(* IEC 61131-3 sources: plcassist-cli/packages/volt-lsp-iec/test-corpus/lenze-mid/Device/Plc Logic/Application/Library Manager/VisuUserManagement, 50 files *)

(* ---- GVL_USERMGMTPROVIDER.gvl ---- *)
VAR_GLOBAL
	G_ARRUSERSTODISPLAY : ARRAY [0..14] OF VUM_UserInternal;
END_VAR

(* ---- VUM_ERRORCODES.gvl ---- *)
VAR_GLOBAL
	ERR_OK : UDINT := 16#0;
	ERR_FAILED : UDINT := 16#1;
	ERR_PARAMETER : UDINT := 16#2;
	ERR_VUM_FILE_NOT_FOUND : UDINT := 16#5000;
	ERR_VUM_TEMP_FILE_CANNOT_BE_OPENED : UDINT := 16#5001;
	ERR_VUM_FILE_READ_FAILED : UDINT := 16#5002;
	ERR_VUM_FILE_WRITE_FAILED : UDINT := 16#5003;
	ERR_VUM_INVALID_FILE_CONTENT : UDINT := 16#5004;
	ERR_VUM_USERNAME_ALREADY_EXIST : UDINT := 16#5005;
	ERR_VUM_WRONG_PASSWORD : UDINT := 16#5006;
	ERR_VUM_UNEQUAL_PASSWORD : UDINT := 16#5007;
	ERR_VUM_NEW_USER_DB_CANNOT_BE_STORED : UDINT := 16#5008;
	ERR_VUM_ONLY_VISIBLE_USERS_CAN_BE_REMOVED : UDINT := 16#5009;
	ERR_VUM_EMPTY_PASSWORD_NOT_ALLOWED : UDINT := 16#500A;
	ERR_VUM_ANOTHER_CLIENT_EDITS_UM : UDINT := 16#500B;
	ERR_VUM_SYSFILE_ERROR : UDINT := 16#500C;
	ERR_VUM_SETNEWUSERDB_FAILED : UDINT := 16#500D;
	ERR_VUM_PROXY_IS_NOT_IN_IDLE_MODE : UDINT := 16#500E;
	ERR_VUM_DATASERVER_ERROR : UDINT := 16#500F;
	ERR_VUM_DATASERVER_ERROR_USERS : UDINT := 16#5010;
	ERR_VUM_MAX_GROUP_LIMIT : UDINT := 16#5011;
	ERR_VUM_USER_DOES_NOT_EXIST : UDINT := 16#5012;
	ERR_VUM_USER_IS_INACTIVE : UDINT := 16#5013;
	ERR_VUM_NO_LOGIN_PROVIDER_AVAILABLE : UDINT := 16#5014;
	ERR_VUM_NO_CLIENT_MEMORY : UDINT := 16#5015;
	ERR_VUM_NO_USER_LOGGED_IN : UDINT := 16#5016;
	ERR_VUM_NO_VALID_USERGROUP_SET : UDINT := 16#5017;
	ERR_VUM_NO_RIGHT_TO_CHANGE_USERS : UDINT := 16#5018;
	ERR_VUM_NO_USER_MANAGEMENT : UDINT := 16#5019;
	ERR_VUM_USER_NOT_IN_USER_GROUP : UDINT := 16#501A;
	ERR_VUM_EXTERNAL_USER_DATABASE_PROVIDER2_NOT_IMPLEMENTED : UDINT := 16#501B;
	ERR_VUM_LOGIN_WRONG_ATTEMPT : UDINT := 16#501C;
	ERR_VUM_LOGIN_SECONDLAST_WRONG_ATTEMPT : UDINT := 16#501D;
	ERR_VUM_LOGIN_LOCKOUT_TEMP : UDINT := 16#501E;
	ERR_VUM_LOGIN_LOCKOUT_COMPLETE : UDINT := 16#501F;
	ERR_VUM_EMPTY_USER_NAME_NOT_ALLOWED : UDINT := 16#5020;
END_VAR

(* ---- VUM_EVENTS.gvl ---- *)
VAR_GLOBAL
	EVT_VISUUSERMGMTGETUSERCOUNT : UDINT := 16#10001;
	EVT_VISUUSERMGMTGETUSERS : UDINT := 16#10002;
	EVT_VISUUSERMGMTCHECKCHANGEUSER : UDINT := 16#10003;
	EVT_VISUUSERMGMTGETSETDB : UDINT := 16#10004;
	CMPID_CMPVISUSERVER : DWORD := 16#57;
END_VAR

(* ---- VUM_GVL.gvl ---- *)
VAR_GLOBAL
	G_VISUUSERMGMT : IVisuUserManagement4;
	G_VISUUSERMGMT2 : IVisuUserManagement4;
	G_VISUUSERMGMTINTERN : IVisuUserMgmt;
	G_STAPPLICATIONNAME : STRING := '';
	G_VUMUSERGROUPNAMES : ARRAY [0..MAX_USER_GROUPS] OF WSTRING;
	G_VUMUSERGROUPMAXINDEX : DWORD;
	G_BUSEVISUUSERMGMTDATASERVER : BOOL;
	G_UDILASTERROR : UDINT;
	G_SILOGINMAXATTEMPTS : SINT := -1;
	G_ILOGINLOCKOUTTIME : INT := -1;
	G_LOGINMAXATTEMPTSENTRIES : VisuUserMgmtFbLoginMaxAttemptsInfoVector;
	G_LOGINLOCKOUTENTRIES : VisuUserMgmtFbLoginLockoutTimeInfoVector;
	G_VISUUSERMANAGERCOMPONENT : STRING := 'VisuUserManager';
	G_VISUUSERMGMTLOGINDIALOGNAME : STRING := 'VUM_Login';
	G_VISUUSERMGMTCHANGEPASSWORDDIALOGNAME : STRING := 'VUM_ChangePassword';
	G_VISUUSERMGMTUSERMANAGEMENTDIALOGNAME : STRING := 'VisuUserManagement.VUM_UserManagementWide';
	G_VISUUSERMGMTRTSBASED : BOOL := FALSE;
	G_VISUUSERMGMTRTSBASEDPATHNAME : WSTRING(256) := "";
END_VAR

(* ---- VUM_GVL_CONSTANT.gvl ---- *)
VAR_GLOBAL
	USERGROUPFLAG_RIGHT_TO_CHANGE_USER : DWORD := 16#1;
	OUTPUT_INFO : INT := 16#1;
	OUTPUT_WARNING : INT := 16#2;
	OUTPUT_ERROR : INT := 16#4;
	OUTPUT_DEBUG : INT := 16#10;
	INVALID_USERGROUP_ID : DWORD := 16#FFFFFFFF;
	INVALID_DB_ID : DWORD := 16#FFFFFFFF;
	INVALID_SELECTION_OR_POS : DWORD := 16#FFFFFFFF;
	COMMENT_CHAR : WORD := 16#23;
	MAX_VISIBLE_USERS : UDINT := 3;
	MAX_USER_GROUPS : UDINT := 255;
	VISU_USER_MGMT_VERSION : DWORD := 0;
	GETSETDB_FLAGS_GETDB : UINT := 16#1;
	GETSETDB_FLAGS_SETDB : UINT := 16#2;
	GETSETDB_FLAGS_SET_RESULT_OK : UINT := 16#4;
	CHECKCHANGEUSER_FLAGS_CHECKLOGIN : UINT := 16#1;
	CHECKCHANGEUSER_FLAGS_CHANGEUSER : UINT := 16#2;
	INVALID_HANDLE : DWORD := 16#FFFFFFFF;
	TIMER_VALUE_LOCKOUT_ADMIN_USER : SINT := 10;
END_VAR

(* ---- VUM_GVL_PROVIDER.gvl ---- *)
VAR_GLOBAL
	G_VISUUSERMGMTPROVIDER : VisuUserMgmtProvider;
	G_BVISUUSERMGMTDIALOGOPEN : BOOL := FALSE;
	G_POPENUSERMGMTORPASSWORDCLIENT : POINTER TO VisuElems.VisuStructClientData;
	G_VISUCHANGEPASSWORDPROVIDER : VisuChangePasswordProvider;
	G_BVISUCHANGEPASSWORDDIALOGOPEN : BOOL := FALSE;
	G_VISUCHANGEPASSWORDPROVIDERMANAGER : Visu_FbChangePasswordProviderManager;
	G_VISULOGINPROVIDERMANAGER : Visu_FbLoginProviderManager;
END_VAR

(* ---- VUM_GVL_RTSUSERMGT.gvl ---- *)
VAR_GLOBAL
	ASSIGNRTSBASEDUSERMGT : VisuAssignRtsBasedUserMgt;
END_VAR

(* ---- IVISUUSERMGMT.itf ---- *)
INTERFACE IVISUUSERMGMT
END_INTERFACE

METHOD CHANGEUSER : BOOL
VAR_INPUT
	DWUSERDB : DWORD;
	PVUMUSER : POINTER TO VUM_User;
	UDIINDEX : UDINT;
	EEDITTYPE : VUM_EditType;
END_VAR
END_METHOD

METHOD CHANGEUSERPASSWORD : BOOL
VAR_INPUT
	DWUSERDB : DWORD;
	WSTUSERNAME : WSTRING;
	WSTNEWPASSWORD : WSTRING;
	WSTOLDPASSWORD : WSTRING;
END_VAR
END_METHOD

METHOD CHECKLOGININTERN : UDINT
VAR_INPUT
	WSTUSERNAME : WSTRING;
	WSTPASSWORD : WSTRING;
END_VAR
VAR_OUTPUT
	WSTFULLNAME : WSTRING;
	DWUSERGROUPID : DWORD;
END_VAR
END_METHOD

METHOD FILLLANGUAGEGROUPNAMES : BOOL
END_METHOD

METHOD GETCURRENTUSER : VUM_User
END_METHOD

METHOD GETGROUPCOUNT : DWORD
END_METHOD

METHOD GETGROUPFROMID : POINTER TO VUM_UserGroup
VAR_INPUT
	DWGROUPID : DWORD;
END_VAR
END_METHOD

METHOD GETGROUPIDFROMINDEX : DWORD
VAR_INPUT
	UDIINDEX : DWORD;
END_VAR
END_METHOD

METHOD GETGROUPINDEXFROMID : DWORD
VAR_INPUT
	DWGROUPID : DWORD;
END_VAR
END_METHOD

METHOD GETLASTERROR : UDINT
END_METHOD

METHOD GETTEXTIDFROMGROUPID : DWORD
VAR_INPUT
	DWGROUPID : DWORD;
END_VAR
END_METHOD

METHOD GETUSERCOUNT : UDINT
VAR_INPUT
	DWUSERDB : DWORD;
END_VAR
END_METHOD

METHOD GETUSERDBASCOPY : DWORD
END_METHOD

METHOD GETUSERS : DWORD
VAR_INPUT
	DWUSERDB : DWORD;
	UDISTARTINDEX : UDINT;
	UDIENDINDEX : UDINT;
	PARR : POINTER TO ARRAY [0..0] OF VUM_User;
	UDIARRSIZE : UDINT;
END_VAR
END_METHOD

METHOD REGISTEREXTERNALUSERDATABASEPROVIDER : VUM_ReturnValues
VAR_INPUT
	ITFEXTENALUSERDATABASEPROVIDER : IExternalUserDatabaseProvider;
END_VAR
END_METHOD

METHOD SETLASTERROR : BOOL
VAR_INPUT
	UDILASTERROR : UDINT;
END_VAR
END_METHOD

METHOD SETNEWUSERDB : BOOL
VAR_INPUT
	DWUSERDB : DWORD;
	BRESULTOK : BOOL;
END_VAR
END_METHOD

METHOD SETPROVIDER : BOOL
VAR_INPUT
	ITFVISUUSERMGMTPROVIDER : IVisuUserMgmtProvider;
END_VAR
END_METHOD

(* ---- IVISUUSERMGMT2.itf ---- *)
INTERFACE IVISUUSERMGMT2
END_INTERFACE

METHOD CHECKTEMPORARYLOCKEDUSER : BOOL
END_METHOD

(* ---- IVISUUSERMGMT3.itf ---- *)
INTERFACE IVISUUSERMGMT3
END_INTERFACE

METHOD CHANGEUSER3 : BOOL
VAR_INPUT
	PCLIENTDATA : POINTER TO VisuElems.VisuStructClientData;
	DWUSERDB : DWORD;
	PVUMUSERNEW : POINTER TO VUM_User;
	PVUMUSEROLD : POINTER TO VUM_User;
	UDIINDEX : UDINT;
	EEDITTYPE : VUM_EditType;
END_VAR
END_METHOD

METHOD CHANGEUSERPASSWORD3 : UDINT
VAR_INPUT
	PCLIENTDATA : POINTER TO VisuElems.VisuStructClientData;
	DWUSERDB : DWORD;
	WSTUSERNAME : WSTRING;
	WSTNEWPASSWORD : WSTRING;
	WSTOLDPASSWORD : WSTRING;
END_VAR
END_METHOD

METHOD CHECKADMINRIGHTS : VUM_UserAdminAccess
VAR_INPUT
	PCLIENTDATA : POINTER TO VisuElems.VisuStructClientData;
END_VAR
END_METHOD

METHOD CHECKGROUPS : BOOL
VAR_INPUT
	PCLIENTDATA : POINTER TO VisuElems.VisuStructClientData;
END_VAR
END_METHOD

METHOD GETUSERCOUNT3 : UDINT
VAR_INPUT
	PCLIENTDATA : POINTER TO VisuElems.VisuStructClientData;
	DWUSERDB : DWORD;
END_VAR
VAR_OUTPUT
	RESULT : RTS_IEC_RESULT;
END_VAR
END_METHOD

METHOD GETUSERS3 : DWORD
VAR_INPUT
	PCLIENTDATA : POINTER TO VisuElems.VisuStructClientData;
	DWUSERDB : DWORD;
	UDISTARTINDEX : UDINT;
	UDIENDINDEX : UDINT;
	PARR : POINTER TO ARRAY [0..0] OF VUM_User;
	UDIARRSIZE : UDINT;
END_VAR
END_METHOD

METHOD LOGINRTS : UDINT
VAR_INPUT
	WSTUSERNAME : WSTRING;
	WSTPASSWORD : WSTRING;
	PCLIENTDATA : POINTER TO VisuElems.VisuStructClientData;
	PUSER : POINTER TO VUM_User;
END_VAR
VAR_OUTPUT
	WSTFULLNAME : WSTRING;
	DWUSERGROUPID : DWORD;
END_VAR
END_METHOD

(* ---- IVISUUSERMGMT4.itf ---- *)
INTERFACE IVISUUSERMGMT4
END_INTERFACE

METHOD CHANGEUSER4 : BOOL
VAR_INPUT
	PCLIENTDATA : POINTER TO VisuElems.VisuStructClientData;
	DWUSERDB : DWORD;
	PVUMUSERNEW : POINTER TO VUM_UserInternal;
	PVUMUSEROLD : POINTER TO VUM_UserInternal;
	UDIINDEX : UDINT;
	EEDITTYPE : VUM_EditType;
END_VAR
END_METHOD

METHOD GETUSERS4 : DWORD
VAR_INPUT
	PCLIENTDATA : POINTER TO VisuElems.VisuStructClientData;
	DWUSERDB : DWORD;
	UDISTARTINDEX : UDINT;
	UDIENDINDEX : UDINT;
	PARR : POINTER TO ARRAY [0..0] OF VUM_UserInternal;
	UDIARRSIZE : UDINT;
END_VAR
END_METHOD

METHOD LOGOUTRTS
VAR_INPUT
	PCLIENTDATA : POINTER TO VisuElems.VisuStructClientData;
END_VAR
END_METHOD

(* ---- IVISUUSERMGMTPROVIDER.itf ---- *)
INTERFACE IVISUUSERMGMTPROVIDER
END_INTERFACE

METHOD SETUSERCOUNT : BOOL
VAR_INPUT
	UDIUSERCOUNT : UDINT;
END_VAR
END_METHOD

METHOD SETUSERDB : BOOL
VAR_INPUT
	UDIUSERDB : UDINT;
END_VAR
END_METHOD

METHOD SETUSERS : BOOL
VAR_INPUT
	UDIUSERCOUNT : UDINT;
	PARRUSERS : POINTER TO ARRAY [0..(MAX_VISIBLE_USERS - 1)] OF VUM_User;
END_VAR
END_METHOD

(* ---- COPYVUM_USER.fun ---- *)
FUNCTION COPYVUM_USER : BOOL
VAR_INPUT
	PVUM_USER : POINTER TO VUM_User;
	PVUM_USERINTERNAL : POINTER TO VUM_UserInternal;
	XFROMUSERTOINTERNAL : BOOL;
END_VAR
END_FUNCTION

(* ---- COPYVUM_USER3.fun ---- *)
FUNCTION COPYVUM_USER3 : BOOL
VAR_INPUT
	PVUM_USER3 : POINTER TO VUM_User3;
	PVUM_USERINTERNAL : POINTER TO VUM_UserInternal;
	XFROMUSERTOINTERNAL : BOOL;
END_VAR
END_FUNCTION

(* ---- FILTERERRORCODE.fun ---- *)
FUNCTION FILTERERRORCODE : UDINT
VAR_INPUT
	ERROR : UDINT;
END_VAR
END_FUNCTION

(* ---- HASUSERGROUPADMINRIGHTS.fun ---- *)
FUNCTION HASUSERGROUPADMINRIGHTS : BOOL
VAR_INPUT
	PUSERGROUP : POINTER TO VUM_UserGroup;
	PCLIENTDATA : POINTER TO VisuElems.VisuStructClientData;
END_VAR
END_FUNCTION

(* ---- ONCHANGEPASSWORDDIALOGCLOSED.fun ---- *)
FUNCTION ONCHANGEPASSWORDDIALOGCLOSED : BOOL
VAR_INPUT
	PCLIENTDATA : POINTER TO VisuElems.VisuStructClientData;
END_VAR
END_FUNCTION

(* ---- ONLOGINDIALOGCLOSED.fun ---- *)
FUNCTION ONLOGINDIALOGCLOSED : BOOL
VAR_INPUT
	PCLIENTDATA : POINTER TO VisuElems.VisuStructClientData;
END_VAR
END_FUNCTION

(* ---- ONUSERMANAGEMENTDIALOGCLOSED.fun ---- *)
FUNCTION ONUSERMANAGEMENTDIALOGCLOSED : BOOL
VAR_INPUT
	PCLIENTDATA : POINTER TO VisuElems.VisuStructClientData;
END_VAR
END_FUNCTION

(* ---- OPENCHANGEPASSWORDDIALOG.fun ---- *)
FUNCTION OPENCHANGEPASSWORDDIALOG : BOOL
VAR_INPUT
	PCLIENTDATA : POINTER TO VisuElems.VisuStructClientData;
END_VAR
END_FUNCTION

(* ---- OPENLOGINDIALOG.fun ---- *)
FUNCTION OPENLOGINDIALOG : BOOL
VAR_INPUT
	PCLIENTDATA : POINTER TO VisuElems.VisuStructClientData;
END_VAR
END_FUNCTION

(* ---- OPENUSERMANAGEMENTDIALOG.fun ---- *)
FUNCTION OPENUSERMANAGEMENTDIALOG : BOOL
VAR_INPUT
	PCLIENTDATA : POINTER TO VisuElems.VisuStructClientData;
END_VAR
END_FUNCTION

(* ---- PRVCHECKUSERMGRISACTIVE.fun ---- *)
FUNCTION PRVCHECKUSERMGRISACTIVE : BOOL
END_FUNCTION

(* ---- SWAPBYTEARRAYBYWORDS.fun ---- *)
FUNCTION SWAPBYTEARRAYBYWORDS : BOOL
VAR_INPUT
	PDATA : POINTER TO ARRAY [0..20] OF BYTE;
	DWSIZE : DWORD;
END_VAR
END_FUNCTION

(* ---- UTILFILLLANGUAGEGROUPNAMES.fun ---- *)
FUNCTION UTILFILLLANGUAGEGROUPNAMES : BOOL
VAR_INPUT
	PARRUSERGROUPTEXTIDS : POINTER TO ARRAY [0..0] OF DWORD;
	DWARRAYSIZE : DWORD;
END_VAR
END_FUNCTION

(* ---- UTILGETFILESIZE.fun ---- *)
FUNCTION UTILGETFILESIZE : UDINT
VAR_INPUT
	DWHANDLE : SysFile.RTS_IEC_HANDLE;
	STFILENAME : REFERENCE TO STRING(255);
	PULRESULT : POINTER TO UDINT;
END_VAR
END_FUNCTION

(* ---- UTILGETMD5HASH.fun ---- *)
FUNCTION UTILGETMD5HASH : BOOL
VAR_INPUT
	PDATA : POINTER TO BYTE;
	DWSIZE : DWORD;
	PMD5HASH : POINTER TO ARRAY [0..15] OF BYTE;
	BADDMAGICNUMBER : BOOL;
	BBYTEORDERMOTOROLAONPOWERPC : BOOL;
END_VAR
END_FUNCTION

(* ---- VISU_FCTINTELBYTEORDER.fun ---- *)
FUNCTION VISU_FCTINTELBYTEORDER : BOOL
END_FUNCTION

(* ---- VISUCREATEUSERMGMTOBJECTS.fun ---- *)
FUNCTION VISUCREATEUSERMGMTOBJECTS : RTS_IEC_RESULT
VAR_INPUT
	PUSERGROUPS : POINTER TO ARRAY [0..0] OF VUM_UserGroup;
	IARRAYSIZE : INT;
	PSAPPNAME : POINTER TO WSTRING;
END_VAR
END_FUNCTION

(* ---- VISUUSERMGMTHASUSERRIGHTTOCHANGEUSERS.fun ---- *)
FUNCTION VISUUSERMGMTHASUSERRIGHTTOCHANGEUSERS : BOOL
VAR_INPUT
	PVUMUSER : POINTER TO VUM_User;
	ITFVISUUSERMGMT : IVisuUserMgmt;
END_VAR
END_FUNCTION

(* ---- VISUUSERMGMTISRTS_GE_35_8.fun ---- *)
FUNCTION VISUUSERMGMTISRTS_GE_35_8 : BOOL
END_FUNCTION

(* ---- VISUUSERMGMTLOG.fun ---- *)
FUNCTION VISUUSERMGMTLOG : BOOL
VAR_INPUT
	DICLASS : DINT;
	DIERROR : DINT;
	DIINFO : DINT;
	STMESSAGE : STRING(255);
END_VAR
END_FUNCTION

(* ---- VISUUSERMGMTSERIALIZEVERSION.fun ---- *)
FUNCTION VISUUSERMGMTSERIALIZEVERSION : DWORD
VAR_INPUT
	VER : VERSION;
END_VAR
END_FUNCTION

(* ---- GLOBALTEXTLIST.fb ---- *)
FUNCTION_BLOCK GLOBALTEXTLIST
VAR
	M_TEXTLISTFILE : STRING(255);
	_STNAMESPACE : STRING;
END_VAR
END_FUNCTION_BLOCK

(* ---- IMAGEPOOL.fb ---- *)
FUNCTION_BLOCK IMAGEPOOL
VAR
	M_STNAMESPACE : STRING(80);
	M_STHELPVARID : STRING;
	M_STHELPVARPATH : STRING(255);
	M_STHELP : STRING;
	M_REGISTERIMAGES : BOOL := TRUE;
END_VAR
END_FUNCTION_BLOCK

METHOD FB_INIT : BOOL
VAR_INPUT
	BINITRETAINS : BOOL;
	BINCOPYCODE : BOOL;
END_VAR
END_METHOD

METHOD FB_REINIT : BOOL
END_METHOD

METHOD FB_EXIT : BOOL
VAR_INPUT
	BINCOPYCODE : BOOL;
END_VAR
END_METHOD

(* ---- IP_VUM.fb ---- *)
FUNCTION_BLOCK IP_VUM
VAR
	M_STNAMESPACE : STRING(80);
	M_STHELPVARID : STRING;
	M_STHELPVARPATH : STRING(255);
	M_STHELP : STRING;
	M_REGISTERIMAGES : BOOL := TRUE;
END_VAR
END_FUNCTION_BLOCK

METHOD FB_INIT : BOOL
VAR_INPUT
	BINITRETAINS : BOOL;
	BINCOPYCODE : BOOL;
END_VAR
END_METHOD

METHOD FB_REINIT : BOOL
END_METHOD

METHOD FB_EXIT : BOOL
VAR_INPUT
	BINCOPYCODE : BOOL;
END_VAR
END_METHOD

(* ---- TL_VUM_ERRORS.fb ---- *)
FUNCTION_BLOCK TL_VUM_ERRORS
VAR
	M_TEXTLISTFILE : STRING(255);
	_STNAMESPACE : STRING;
END_VAR
END_FUNCTION_BLOCK

(* ---- VISU_FBCHANGEPASSWORDPROVIDERMANAGER.fb ---- *)
FUNCTION_BLOCK VISU_FBCHANGEPASSWORDPROVIDERMANAGER
VAR
	M_ARRPROVIDER : ARRAY [0..(MAX_PROVIDER - 1)] OF VisuChangePasswordProvider;
	M_ARRCLIENT : ARRAY [0..(MAX_PROVIDER - 1)] OF POINTER TO VisuElems.VisuStructClientData;
	M_ITFCLIENTMANAGERLISTENER : VisuElems.IClientManagerListener := THIS^;
	M_BINIT : BOOL;
	I : INT;
	MAX_PROVIDER : INT := 5;
END_VAR
END_FUNCTION_BLOCK

METHOD FB_EXIT : BOOL
VAR_INPUT
	BINCOPYCODE : BOOL;
END_VAR
END_METHOD

METHOD INITIALIZE : BOOL
END_METHOD

METHOD REGISTERCLIENT : POINTER TO VisuChangePasswordProvider
VAR_INPUT
	PCLIENTDATA : POINTER TO VisuElems.VisuStructClientData;
END_VAR
END_METHOD

METHOD UNREGISTERCLIENT : BOOL
VAR_INPUT
	PCLIENTDATA : POINTER TO VisuElems.VisuStructClientData;
END_VAR
END_METHOD

METHOD CLIENTCREATED
VAR_INPUT
	PCLIENTDATA : POINTER TO VisuElems.VisuStructClientData;
END_VAR
END_METHOD

METHOD CLIENTDESTROYED
VAR_INPUT
	PCLIENTDATA : POINTER TO VisuElems.VisuStructClientData;
END_VAR
END_METHOD

(* ---- VISU_FBLOGINPROVIDERMANAGER.fb ---- *)
FUNCTION_BLOCK VISU_FBLOGINPROVIDERMANAGER
VAR
	M_ARRLOGINPROVIDER : ARRAY [0..(MAX_LOGIN_PROVIDER - 1)] OF VisuLoginProvider;
	M_ARRLOGINPROVIDERSET : ARRAY [0..(MAX_LOGIN_PROVIDER - 1)] OF BOOL;
	M_ITFCLIENTMANAGERLISTENER : VisuElems.IClientManagerListener := THIS^;
	M_BINIT : BOOL;
	I : INT;
	MAX_LOGIN_PROVIDER : INT := 5;
END_VAR
END_FUNCTION_BLOCK

METHOD FB_EXIT : BOOL
VAR_INPUT
	BINCOPYCODE : BOOL;
END_VAR
END_METHOD

METHOD INITIALIZE : BOOL
END_METHOD

METHOD REGISTERLOGINPROVIDERCLIENT : POINTER TO VisuLoginProvider
VAR_INPUT
	PCLIENTDATA : POINTER TO VisuElems.VisuStructClientData;
END_VAR
END_METHOD

METHOD UNREGISTERLOGINPROVIDERCLIENT : BOOL
VAR_INPUT
	PCLIENTDATA : POINTER TO VisuElems.VisuStructClientData;
END_VAR
END_METHOD

METHOD CLIENTCREATED
VAR_INPUT
	PCLIENTDATA : POINTER TO VisuElems.VisuStructClientData;
END_VAR
END_METHOD

METHOD CLIENTDESTROYED
VAR_INPUT
	PCLIENTDATA : POINTER TO VisuElems.VisuStructClientData;
END_VAR
END_METHOD

(* ---- VISUASSIGNRTSBASEDUSERMGT.fb ---- *)
FUNCTION_BLOCK VISUASSIGNRTSBASEDUSERMGT
VAR
	XSTATUSVISUUSERMGMTRTSBASED : BOOL;
END_VAR
END_FUNCTION_BLOCK

METHOD FB_EXIT : BOOL
VAR_INPUT
	BINCOPYCODE : BOOL;
END_VAR
END_METHOD

METHOD FB_INIT : BOOL
VAR_INPUT
	BINITRETAINS : BOOL;
	BINCOPYCODE : BOOL;
END_VAR
END_METHOD

(* ---- VISUCHANGEPASSWORDPROVIDER.fb ---- *)
FUNCTION_BLOCK VISUCHANGEPASSWORDPROVIDER
VAR
	STUSERNAME : WSTRING;
	STOLDPASSWORD : WSTRING;
	STPASSWORD : WSTRING;
	WSTOLDPASSWORD : WSTRING;
	STACKNOWLEDGEPASSWORD : WSTRING;
	DWDIALOGRESULTOK : BOOL;
	DWLASTDIALOGRESULTOK : BOOL;
	DWDIALOGRESULTCANCEL : BOOL;
	DWLASTDIALOGRESULTCANCEL : BOOL;
	UDILASTERROR : UDINT;
	DWRESULT : DWORD;
	VUMUSER : VUM_User;
	BRTSBASED : BOOL;
	BCHGPASSWORD : BOOL;
	_IVISUUSERMGMT : IVisuUserMgmt;
	_IVISUUSERMGMT4 : IVisuUserMgmt4;
	_VISUUSERMGMTSTATE : EVisuUserMgmtState;
	_PCLIENTDATA : POINTER TO VisuElems.VisuStructClientData;
	_BCURRENTSTATE : BYTE := 0;
	_BLASTCURRENTSTATE : BYTE := 0;
	_DWUSERDB : DWORD;
	VCPP_STATE_NONE : BYTE := 0;
	VCPP_STATE_GET_USER_DB : BYTE := 1;
	VCPP_STATE_CHECK_LOGIN : BYTE := 2;
	VCPP_STATE_CHANGE_USER_PASSWORD : BYTE := 3;
	VCPP_STATE_SET_USER_DB : BYTE := 4;
END_VAR
END_FUNCTION_BLOCK

METHOD CHECKPASSWORD : BOOL
END_METHOD

METHOD INITIALIZE : BOOL
VAR_INPUT
	IVISUUSERMGMT : IVisuUserMgmt;
	PCLIENTDATA : POINTER TO VisuElems.VisuStructClientData;
END_VAR
END_METHOD

METHOD SETUSERCOUNT : BOOL
VAR_INPUT
	UDIUSERCOUNT : UDINT;
END_VAR
END_METHOD

METHOD SETUSERDB : BOOL
VAR_INPUT
	UDIUSERDB : UDINT;
END_VAR
END_METHOD

METHOD SETUSERS : BOOL
VAR_INPUT
	UDIUSERCOUNT : UDINT;
	PARRUSERS : POINTER TO ARRAY [0..(MAX_VISIBLE_USERS - 1)] OF VUM_User;
END_VAR
END_METHOD

METHOD PRVFILLUSER : BOOL
END_METHOD

METHOD PRVSETNEWUSERDB : BOOL
VAR_INPUT
	DWUSERDB : DWORD;
	BRESULTOK : BOOL;
END_VAR
END_METHOD

(* ---- VISUFBCLIENTMANAGERLISTENER.fb ---- *)
FUNCTION_BLOCK VISUFBCLIENTMANAGERLISTENER
END_FUNCTION_BLOCK

METHOD CLIENTCREATED
VAR_INPUT
	PCLIENTDATA : POINTER TO VisuElems.VisuStructClientData;
END_VAR
END_METHOD

METHOD CLIENTDESTROYED
VAR_INPUT
	PCLIENTDATA : POINTER TO VisuElems.VisuStructClientData;
END_VAR
END_METHOD

(* ---- VISULOGINPROVIDER.fb ---- *)
FUNCTION_BLOCK VISULOGINPROVIDER
VAR
	STUSERNAME : WSTRING;
	STPASSWORD : WSTRING;
	DWDIALOGRESULTOK : BOOL;
	DWLASTDIALOGRESULTOK : BOOL;
	DWDIALOGRESULTCANCEL : BOOL;
	DWLASTDIALOGRESULTCANCEL : BOOL;
	UDILASTERROR : UDINT;
	VUMUSER : VUM_User;
	BRTSBASED : BOOL;
	_IVISUUSERMGMT : IVisuUserMgmt;
	_IVISUUSERMGMT3 : IVisuUserMgmt3;
	_VISUUSERMGMTSTATE : EVisuUserMgmtState;
	_VUMCURRENTUSER : VUM_User;
	_PCLIENTDATA : POINTER TO VisuElems.VisuStructClientData;
	_BCURRENTSTATE : BYTE := 0;
	_BLASTCURRENTSTATE : BYTE := 0;
	_DWUSERGROUPID : DWORD;
	_XDOIT : BOOL;
	_DWPROP : DWORD;
	_SUSER : STRING;
	_RESULT : RTS_IEC_RESULT;
	VLP_STATE_NONE : BYTE := 0;
	VLP_STATE_CHECK_LOGIN : BYTE := 2;
END_VAR
END_FUNCTION_BLOCK

METHOD CHECKLOGIN : BOOL
END_METHOD

METHOD DELETELOGINATTEMPTSINFOS : BOOL
VAR_INPUT
	WSTUSERNAMETODELETE : WSTRING;
END_VAR
END_METHOD

METHOD INITIALIZE : BOOL
VAR_INPUT
	IVISUUSERMGMT : IVisuUserMgmt;
	PCLIENTDATA : POINTER TO VisuElems.VisuStructClientData;
END_VAR
END_METHOD

METHOD LOGIN : UDINT
VAR_OUTPUT
	WSTFULLNAME : WSTRING;
	DWUSERGROUPID : DWORD;
	ABYUSERGROUPIDS : ARRAY [0..VUM_Constants.VISU_VUM_MAX_GROUPS_PER_USER] OF BYTE;
	BYUSERGROUPCOUNT : BYTE;
	BDEACTIVATED : BOOL;
END_VAR
END_METHOD

METHOD UPDATELOGINATTEMPTSINFOS : BOOL
VAR_INPUT
	LASTATTEMPTSTATE : UDINT;
END_VAR
END_METHOD

METHOD SETLASTRESULT : BOOL
VAR_INPUT
	UDILASTRESULT : UDINT;
END_VAR
END_METHOD

METHOD SETUSERCOUNT : BOOL
VAR_INPUT
	UDIUSERCOUNT : UDINT;
END_VAR
END_METHOD

METHOD SETUSERDB : BOOL
VAR_INPUT
	UDIUSERDB : UDINT;
END_VAR
END_METHOD

METHOD SETUSERS : BOOL
VAR_INPUT
	UDIUSERCOUNT : UDINT;
	PARRUSERS : POINTER TO ARRAY [0..(MAX_VISIBLE_USERS - 1)] OF VUM_User;
END_VAR
END_METHOD

METHOD PRVCHECKCURRENTUSERISADMIN : BOOL
VAR_INPUT
	DWCURRENTUSERDBCOPY : DWORD;
END_VAR
END_METHOD

METHOD PRVGETTIMESTAMPINMINUTES
VAR_OUTPUT
	DWTIMESTAMP : DWORD;
END_VAR
END_METHOD

METHOD PRVGETUSERANDINDEXBYNAME : BOOL
VAR_INPUT
	WSTUSERNAMETOFIND : WSTRING;
END_VAR
VAR_OUTPUT
	VUMUSERFOUND : VUM_User;
	UDIUSERINDEX : UDINT;
END_VAR
END_METHOD

METHOD PRVLOGIN : BOOL
VAR_INPUT
	XCOMPLETEEXEC : BOOL;
END_VAR
END_METHOD

(* ---- VISUUSERMGMT.fb ---- *)
FUNCTION_BLOCK VISUUSERMGMT
VAR
	_PARRUSERGROUPS : POINTER TO ARRAY [0..0] OF VUM_UserGroup;
	_PARRUSERGROUPTEXTIDS : POINTER TO ARRAY [0..0] OF DWORD;
	_DWARRAYSIZE : DWORD := 0;
	_UDILASTERROR : UDINT := 0;
	_UDILASTRESULT : UDINT := 0;
	_UDILASTFILEERROR : UDINT := 0;
	_STLASTFILEERRORPOS : STRING := '';
	_STSEPARATOR : WSTRING(1) := ";";
	_STPIPESEPARATOR : WSTRING(1) := "|";
	_STNEWLINE : WSTRING(2) := "$R$N";
	_WUNICODEFILE : WORD := 16#FEFF;
	_BUNICODEFILE1 : BYTE := 16#FF;
	_BUNICODEFILE2 : BYTE := 16#FE;
	_VUMCURRENTUSER : VUM_User;
	_DATABUFFER : ARRAY [0..MAX_BUFFER_SIZE] OF BYTE;
	_CURRENTDATAPOSITION : DWORD;
	_BNOSYSFILEWRITEHAPPEND : BOOL;
	_DWNEXTUSERDB : DWORD := 1;
	_ARRERRORQUEUE : ARRAY [0..20] OF UDINT;
	_ITFEXTERNALUSERDATABASEPROVIDER : IExternalUserDatabaseProvider;
	_BCHECKUSERWITHTEMPLOCKOUT : BOOL;
	_ICURRENTUSERLOCKOUTTIME : INT := -1;
	_TONINST : TON;
	_BTIMEOFF : BOOL;
	_BSTARTTIMER : BOOL;
	_ITIMER : INT;
	MAX_ERRORS : INT := 20;
	MAX_BUFFER_SIZE : DWORD := 4000;
	USER_MANAGEMENT_FILE_NAME : STRING := 'visuusermgmtdb';
	USER_MANAGEMENT_STORAGE_VERSION : WSTRING := "V1.0.0.0";
	LOGIN_TYPE_CHECK : INT := 0;
	LOGIN_TYPE_LOGIN : INT := 1;
	LOGIN_TYPE_RELOGIN : INT := 2;
	S_SEM : VisuUserMgmtSem;
	CHECKUSERWITHTEMPLOCKOUT : BOOL;
	CURRENTUSERLOCKOUTTIME : INT;
	LASTRESULT : UDINT;
	STATE : EVisuUserMgmtState;
END_VAR
END_FUNCTION_BLOCK

METHOD CHANGELANGUAGE : BOOL
END_METHOD

METHOD CHANGEUSER : BOOL
VAR_INPUT
	DWUSERDB : DWORD;
	PVUMUSER : POINTER TO VUM_User;
	UDIINDEX : UDINT;
	EEDITTYPE : VUM_EditType;
END_VAR
END_METHOD

METHOD CHANGEUSERPASSWORD : BOOL
VAR_INPUT
	DWUSERDB : DWORD;
	WSTUSERNAME : WSTRING;
	WSTNEWPASSWORD : WSTRING;
	WSTOLDPASSWORD : WSTRING;
END_VAR
END_METHOD

METHOD CHECKLOGININTERN : UDINT
VAR_INPUT
	WSTUSERNAME : WSTRING;
	WSTPASSWORD : WSTRING;
END_VAR
VAR_OUTPUT
	WSTFULLNAME : WSTRING;
	DWUSERGROUPID : DWORD;
END_VAR
END_METHOD

METHOD CHECKLOGINWITHGROUPIDINTERN : UDINT
VAR_INPUT
	WSTUSERNAME : WSTRING;
	WSTPASSWORD : WSTRING;
	DWUSERGROUPID : DWORD;
END_VAR
VAR_OUTPUT
	WSTFULLNAME : WSTRING;
END_VAR
END_METHOD

METHOD FB_INIT : BOOL
VAR_INPUT
	BINITRETAINS : BOOL;
	BINCOPYCODE : BOOL;
END_VAR
END_METHOD

METHOD FILLLANGUAGEGROUPNAMES : BOOL
END_METHOD

METHOD FINDUSERBYTYPE : VUM_ReturnValues
VAR_INPUT
	VUMUSERIN : VUM_User;
	EEDITTYPE : VUM_EditType;
END_VAR
VAR_OUTPUT
	VUMUSER : VUM_User;
	UDIINDEX : UDINT;
END_VAR
END_METHOD

METHOD GETCURRENTUSER : VUM_User
END_METHOD

METHOD GETGROUPCOUNT : DWORD
END_METHOD

METHOD GETGROUPFROMID : POINTER TO VUM_UserGroup
VAR_INPUT
	DWGROUPID : DWORD;
END_VAR
END_METHOD

METHOD GETGROUPIDFROMINDEX : DWORD
VAR_INPUT
	UDIINDEX : DWORD;
END_VAR
END_METHOD

METHOD GETGROUPINDEXFROMID : DWORD
VAR_INPUT
	DWGROUPID : DWORD;
END_VAR
END_METHOD

METHOD GETGROUPNAMEFROMID : WSTRING
VAR_INPUT
	DWGROUPID : DWORD;
END_VAR
END_METHOD

METHOD GETLASTERROR : UDINT
END_METHOD

METHOD GETTEXTIDFROMGROUPID : DWORD
VAR_INPUT
	DWGROUPID : DWORD;
END_VAR
END_METHOD

METHOD GETUSERCOUNT : UDINT
VAR_INPUT
	DWUSERDB : DWORD;
END_VAR
END_METHOD

METHOD GETUSERDBASCOPY : DWORD
END_METHOD

METHOD GETUSERS : DWORD
VAR_INPUT
	DWUSERDB : DWORD;
	UDISTARTINDEX : UDINT;
	UDIENDINDEX : UDINT;
	PARR : POINTER TO ARRAY [0..0] OF VUM_User;
	UDIARRSIZE : UDINT;
END_VAR
END_METHOD

METHOD INITIALIZE : BOOL
VAR_INPUT
	PARRUSERGROUPS : POINTER TO ARRAY [0..0] OF VUM_UserGroup;
	PARRUSERGROUPTEXTIDS : POINTER TO ARRAY [0..0] OF DWORD;
	DWARRAYSIZE : DWORD;
END_VAR
END_METHOD

METHOD SETLASTERROR : BOOL
VAR_INPUT
	UDILASTERROR : UDINT;
END_VAR
END_METHOD

METHOD SETNEWUSERDB : BOOL
VAR_INPUT
	DWUSERDB : DWORD;
	BRESULTOK : BOOL;
END_VAR
END_METHOD

METHOD LOGOUTUSER : DWORD
VAR_INPUT
	PCLIENTDATA : POINTER TO VisuElems.VisuStructClientData;
END_VAR
END_METHOD

METHOD NEWSESSION : DWORD
VAR_INPUT
	PCLIENTDATA : POINTER TO VisuElems.VisuStructClientData;
	DWSESSIONID : DWORD;
END_VAR
END_METHOD

METHOD CHECKLOGINWITHGROUPID : VUM_ReturnValues
VAR_INPUT
	WSTUSERNAME : WSTRING;
	WSTPASSWORD : WSTRING;
	DWUSERGROUPID : DWORD;
END_VAR
END_METHOD

METHOD CHECKLOGIN : VUM_ReturnValues
VAR_INPUT
	WSTUSERNAME : WSTRING;
	WSTPASSWORD : WSTRING;
END_VAR
END_METHOD

METHOD REGISTEREXTERNALUSERDATABASEPROVIDER : VUM_ReturnValues
VAR_INPUT
	ITFEXTENALUSERDATABASEPROVIDER : IExternalUserDatabaseProvider;
END_VAR
END_METHOD

METHOD LOGINTOUSERGROUP : BOOL
VAR_INPUT
	PCLIENT : POINTER TO BYTE;
	DWGROUPID : DWORD;
	WSTUSERNAME : WSTRING(79);
	WSTFULLNAME : WSTRING(79);
END_VAR
END_METHOD

METHOD LOGINTOUSERGROUPS : BOOL
VAR_INPUT
	PCLIENT : POINTER TO BYTE;
	PADWUSERGROUPIDS : POINTER TO ARRAY [0..0] OF DWORD;
	DWUSERGROUPCOUNT : DWORD;
	WSTUSERNAME : WSTRING(79);
	WSTFULLNAME : WSTRING(79);
END_VAR
END_METHOD

METHOD CHANGEPASSWORD : VUM_ReturnValues
VAR_INPUT
	PCLIENT : POINTER TO BYTE;
	WSTUSERNAME : WSTRING(79);
	WSTNEWPASSWORD : WSTRING(79);
	WSTOLDPASSWORD : WSTRING(79);
END_VAR
END_METHOD

METHOD LOGIN : VUM_ReturnValues
VAR_INPUT
	PCLIENT : POINTER TO BYTE;
	WSTUSERNAME : WSTRING(79);
	WSTPASSWORD : WSTRING(79);
END_VAR
VAR_OUTPUT
	WSTFULLNAMEIFAVAILABLE : WSTRING;
	DWUSERGROUPID : DWORD;
	ADWUSERGROUPIDS : ARRAY [0..VUM_Constants.VISU_VUM_MAX_GROUPS_PER_USER] OF DWORD;
	DWUSERGROUPCOUNT : DWORD;
	BDEACTIVATED : BOOL;
END_VAR
END_METHOD

METHOD LOGOUT : VUM_ReturnValues
VAR_INPUT
	PCLIENT : POINTER TO BYTE;
END_VAR
END_METHOD

METHOD USERCOUNT : UDINT
VAR_INPUT
	PCLIENT : POINTER TO BYTE;
END_VAR
VAR_OUTPUT
	RESULT : VUM_ReturnValues;
END_VAR
END_METHOD

METHOD USERS : VUM_ReturnValues
VAR_INPUT
	PCLIENT : POINTER TO BYTE;
	UDISTARTINDEX : UDINT;
	UDIENDINDEX : UDINT;
	PARR : POINTER TO ARRAY [0..0] OF VUM_User2;
	UDIARRSIZE : UDINT;
END_VAR
END_METHOD

METHOD EDITUSER : VUM_ReturnValues
VAR_INPUT
	PCLIENT : POINTER TO BYTE;
	PVUMUSERNEW : POINTER TO VUM_User3;
	PVUMUSEROLD : POINTER TO VUM_User3;
	UDIINDEX : UDINT;
	EEDITTYPE : VUM_EditType;
END_VAR
END_METHOD

METHOD SETPROVIDER : BOOL
VAR_INPUT
	ITFVISUUSERMGMTPROVIDER : IVisuUserMgmtProvider;
END_VAR
END_METHOD

METHOD CHECKTEMPORARYLOCKEDUSER : BOOL
END_METHOD

METHOD CHANGEUSER3 : BOOL
VAR_INPUT
	PCLIENTDATA : POINTER TO VisuElems.VisuStructClientData;
	DWUSERDB : DWORD;
	PVUMUSERNEW : POINTER TO VUM_User;
	PVUMUSEROLD : POINTER TO VUM_User;
	UDIINDEX : UDINT;
	EEDITTYPE : VUM_EditType;
END_VAR
END_METHOD

METHOD CHANGEUSERPASSWORD3 : UDINT
VAR_INPUT
	PCLIENTDATA : POINTER TO VisuElems.VisuStructClientData;
	DWUSERDB : DWORD;
	WSTUSERNAME : WSTRING;
	WSTNEWPASSWORD : WSTRING;
	WSTOLDPASSWORD : WSTRING;
END_VAR
END_METHOD

METHOD CHECKADMINRIGHTS : VUM_UserAdminAccess
VAR_INPUT
	PCLIENTDATA : POINTER TO VisuElems.VisuStructClientData;
END_VAR
END_METHOD

METHOD CHECKGROUPS : BOOL
VAR_INPUT
	PCLIENTDATA : POINTER TO VisuElems.VisuStructClientData;
END_VAR
END_METHOD

METHOD GETUSERCOUNT3 : UDINT
VAR_INPUT
	PCLIENTDATA : POINTER TO VisuElems.VisuStructClientData;
	DWUSERDB : DWORD;
END_VAR
VAR_OUTPUT
	RESULT : RTS_IEC_RESULT;
END_VAR
END_METHOD

METHOD GETUSERS3 : DWORD
VAR_INPUT
	PCLIENTDATA : POINTER TO VisuElems.VisuStructClientData;
	DWUSERDB : DWORD;
	UDISTARTINDEX : UDINT;
	UDIENDINDEX : UDINT;
	PARR : POINTER TO ARRAY [0..0] OF VUM_User;
	UDIARRSIZE : UDINT;
END_VAR
END_METHOD

METHOD LOGINRTS : UDINT
VAR_INPUT
	WSTUSERNAME : WSTRING;
	WSTPASSWORD : WSTRING;
	PCLIENTDATA : POINTER TO VisuElems.VisuStructClientData;
	PUSER : POINTER TO VUM_User;
END_VAR
VAR_OUTPUT
	WSTFULLNAME : WSTRING;
	DWUSERGROUPID : DWORD;
END_VAR
END_METHOD

METHOD CHANGEUSER4 : BOOL
VAR_INPUT
	PCLIENTDATA : POINTER TO VisuElems.VisuStructClientData;
	DWUSERDB : DWORD;
	PVUMUSERNEW : POINTER TO VUM_UserInternal;
	PVUMUSEROLD : POINTER TO VUM_UserInternal;
	UDIINDEX : UDINT;
	EEDITTYPE : VUM_EditType;
END_VAR
END_METHOD

METHOD GETUSERS4 : DWORD
VAR_INPUT
	PCLIENTDATA : POINTER TO VisuElems.VisuStructClientData;
	DWUSERDB : DWORD;
	UDISTARTINDEX : UDINT;
	UDIENDINDEX : UDINT;
	PARR : POINTER TO ARRAY [0..0] OF VUM_UserInternal;
	UDIARRSIZE : UDINT;
END_VAR
END_METHOD

METHOD LOGOUTRTS
VAR_INPUT
	PCLIENTDATA : POINTER TO VisuElems.VisuStructClientData;
END_VAR
END_METHOD

METHOD PRVCHANGEUSERPASSWORDRTS : DWORD
VAR_INPUT
	PCLIENTDATA : POINTER TO VisuElems.VisuStructClientData;
	WSTUSERNAME : WSTRING;
	WSTNEWPASSWORD : WSTRING;
	WSTOLDPASSWORD : WSTRING;
END_VAR
END_METHOD

METHOD PRVCHANGEUSERRTS : DWORD
VAR_INPUT
	PCLIENTDATA : POINTER TO VisuElems.VisuStructClientData;
	PVUMUSERNEW : POINTER TO VUM_UserInternal;
	PVUMUSEROLD : POINTER TO VUM_UserInternal;
	EEDITTYPE : VUM_EditType;
END_VAR
END_METHOD

METHOD PRVCHANGEUSERRTS_ADD : DWORD
VAR_INPUT
	HUSER : RTS_IEC_HANDLE;
	PVUMUSER : POINTER TO VUM_UserInternal;
END_VAR
END_METHOD

METHOD PRVCHANGEUSERRTS_GRPADD : DWORD
VAR_INPUT
	HUSER : RTS_IEC_HANDLE;
	PVUMUSER : POINTER TO VUM_UserInternal;
END_VAR
END_METHOD

METHOD PRVCHANGEUSERRTS_GRPREMOVE : DWORD
VAR_INPUT
	HUSER : RTS_IEC_HANDLE;
	PVUMUSER : POINTER TO VUM_UserInternal;
END_VAR
END_METHOD

METHOD PRVCHANGEUSERRTS_MODIFY : DWORD
VAR_INPUT
	HUSER : RTS_IEC_HANDLE;
	PVUMUSERNEW : POINTER TO VUM_UserInternal;
	PVUMUSEROLD : POINTER TO VUM_UserInternal;
END_VAR
END_METHOD

METHOD PRVCHANGEUSERRTS_REMOVE : DWORD
VAR_INPUT
	HUSER : RTS_IEC_HANDLE;
	PVUMUSER : POINTER TO VUM_UserInternal;
END_VAR
END_METHOD

METHOD PRVCHECKUSERISADMIN : VUM_UserAdminAccess
VAR_INPUT
	PCLIENTDATA : POINTER TO VisuElems.VisuStructClientData;
END_VAR
END_METHOD

METHOD PRVCONVERTUTF8TOWS : WSTRING(512)
VAR_INPUT
	SORIGINAL : STRING(512);
END_VAR
END_METHOD

METHOD PRVCONVERTWSTOUTF8 : STRING(512)
VAR_INPUT
	WSORIGINAL : WSTRING(512);
END_VAR
END_METHOD

METHOD PRVGETMAPPEDGROUP : DWORD
VAR_INPUT
	HUSER : RTS_IEC_HANDLE;
	WSVISUGRPNAME : WSTRING;
END_VAR
VAR_OUTPUT
	WSMAPPEDGROUP : WSTRING;
END_VAR
END_METHOD

METHOD PRVGETUSERCOUNTRTS : UDINT
VAR_INPUT
	PCLIENTDATA : POINTER TO VisuElems.VisuStructClientData;
END_VAR
VAR_OUTPUT
	RESULT : RTS_IEC_RESULT;
END_VAR
END_METHOD

METHOD PRVGETUSERGROUPSIDS
VAR_INPUT
	HUSER : RTS_IEC_HANDLE;
	PUSER : POINTER TO VUM_UserInternal;
	BRIGHTS : BOOL;
	WSUSERNAME : WSTRING;
END_VAR
END_METHOD

METHOD PRVGETUSERSRTS : DWORD
VAR_INPUT
	PCLIENTDATA : POINTER TO VisuElems.VisuStructClientData;
	UDISTARTINDEX : UDINT;
	UDIENDINDEX : UDINT;
	PARR : POINTER TO ARRAY [0..10] OF VUM_UserInternal;
	UDIARRSIZE : UDINT;
END_VAR
END_METHOD

METHOD PRVISUSERBELONGGROUP : BOOL
VAR_INPUT
	HUSER : RTS_IEC_HANDLE;
	DWUSERGROUPID : DWORD;
END_VAR
END_METHOD

METHOD PRVISUSERBELONGGROUP2 : BOOL
VAR_INPUT
	HUSER : RTS_IEC_HANDLE;
	WSUSERNAME : WSTRING;
	DWUSERGROUPID : DWORD;
END_VAR
END_METHOD

METHOD PRVLOGINBYSESSIONID : DWORD
VAR_INPUT
	PCLIENTDATA : POINTER TO VisuElems.VisuStructClientData;
	DWSESSIONID : DWORD;
END_VAR
END_METHOD

METHOD PRVLOGINRTS
VAR_INPUT
	WSTUSERNAME : WSTRING;
	WSTPASSWORD : WSTRING;
	PCLIENTDATA : POINTER TO VisuElems.VisuStructClientData;
	PUSER : POINTER TO VUM_UserInternal;
	ITYPE : INT;
END_VAR
VAR_OUTPUT
	WSTFULLNAME : WSTRING;
	DWUSERGROUPID : DWORD;
END_VAR
END_METHOD

METHOD PRVLOGINWITHGROUPIDRTS
VAR_INPUT
	WSTUSERNAME : WSTRING;
	WSTPASSWORD : WSTRING;
	DWUSERGROUPID : DWORD;
	PCLIENTDATA : POINTER TO VisuElems.VisuStructClientData;
	XCHECKONLY : BOOL;
END_VAR
VAR_OUTPUT
	WSTFULLNAME : WSTRING;
END_VAR
END_METHOD

METHOD PRVLOGOUTRTS
VAR_INPUT
	PCLIENT : POINTER TO VisuElems.VisuStructClientData;
END_VAR
END_METHOD

METHOD PRVCHECKTEMPORARYLOCKEDUSER : BOOL
END_METHOD

METHOD PRVCHECKUSER : BOOL
VAR_INPUT
	PWORDDATA : POINTER TO WORD;
	PVUMUSER : POINTER TO VUM_User;
	PSTART : POINTER TO DWORD;
	ULSIZE : DWORD;
	PBUSERFOUND : POINTER TO BOOL;
	EEDITTYPE : VUM_EditType;
END_VAR
END_METHOD

METHOD PRVCLEANUSERGROUPSIDS
VAR_INPUT
	PUSER : POINTER TO VUM_User;
END_VAR
END_METHOD

METHOD PRVDELETELOGINATTEMPTSINFOS : BOOL
VAR_INPUT
	WSTUSERNAMETODELETE : WSTRING;
END_VAR
END_METHOD

METHOD PRVFREERESOURCES : BOOL
VAR_INPUT
	PDATA : POINTER TO BYTE;
	DWHANDLE1 : SysFile.RTS_IEC_HANDLE;
	DWHANDLE2 : SysFile.RTS_IEC_HANDLE;
	BSEMLEAVE : BOOL;
END_VAR
END_METHOD

METHOD PRVGETFILENAME : BOOL
VAR_INPUT
	PSTFILENAME : POINTER TO STRING(255);
	DWUSERDB : DWORD;
	BTEMP : BOOL;
END_VAR
END_METHOD

METHOD PRVGETGROUPFROMINDEX : POINTER TO VUM_UserGroup
VAR_INPUT
	IINDEX : DWORD;
END_VAR
END_METHOD

METHOD PRVGETHASHASWSTRING : BOOL
VAR_INPUT
	PSTR : POINTER TO WSTRING(40);
	PHASH : POINTER TO ARRAY [0..15] OF BYTE;
END_VAR
END_METHOD

METHOD PRVGETHASHFROMWSTRING : BOOL
VAR_INPUT
	PSTR : POINTER TO WSTRING(40);
	PHASH : POINTER TO ARRAY [0..15] OF BYTE;
END_VAR
END_METHOD

METHOD PRVGETTIMESTAMPINMINUTES
VAR_OUTPUT
	DWTIMESTAMP : DWORD;
END_VAR
END_METHOD

METHOD PRVMODIFYUSER : BOOL
VAR_INPUT
	DWUSERDB : DWORD;
	PVUMUSER : POINTER TO VUM_User;
	UDIINDEX : UDINT;
	EEDITTYPE : VUM_EditType;
END_VAR
END_METHOD

METHOD PRVREADLINE : POINTER TO WORD
VAR_INPUT
	PDATA : POINTER TO WORD;
	PULSTART : POINTER TO DWORD;
	ULSIZE : DWORD;
END_VAR
END_METHOD

METHOD PRVREADTOKEN : POINTER TO BYTE
VAR_INPUT
	PDATA : POINTER TO WORD;
	PULSTART : POINTER TO DWORD;
	ULSIZE : DWORD;
END_VAR
END_METHOD

METHOD PRVREADUSER : BOOL
VAR_INPUT
	PWORDDATA : POINTER TO WORD;
	PVUMUSER : POINTER TO VUM_User;
	PSTART : POINTER TO DWORD;
	ULSIZE : DWORD;
END_VAR
END_METHOD

METHOD PRVREADUSERGROUP : BOOL
VAR_INPUT
	PVUMUSER : POINTER TO VUM_User;
	PWST : POINTER TO WSTRING;
END_VAR
END_METHOD

METHOD PRVREADUSERS : BOOL
VAR_INPUT
	DWUSERDB : DWORD;
	UDISTARTINDEX : UDINT;
	UDIENDINDEX : UDINT;
	PARR : POINTER TO ARRAY [0..0] OF VUM_User;
	UDIARRSIZE : UDINT;
	PDIUSERCOUNT : POINTER TO DINT;
	BFINDUSER : BOOL;
	EEDITTYPE : VUM_EditType;
END_VAR
END_METHOD

METHOD PRVREADUSERS2 : BOOL
VAR_INPUT
	DWUSERDB : DWORD;
	UDISTARTINDEX : UDINT;
	UDIENDINDEX : UDINT;
	PARR : POINTER TO ARRAY [0..0] OF VUM_User;
	UDIARRSIZE : UDINT;
	PDIUSERCOUNT : POINTER TO DINT;
	BFINDUSER : BOOL;
	EEDITTYPE : VUM_EditType;
END_VAR
VAR_OUTPUT
	VUMUSER : VUM_User;
	UDIINDEX : UDINT;
END_VAR
END_METHOD

METHOD PRVWRITEFILECHECKSUM : BOOL
VAR_INPUT
	PSTFILENAME : POINTER TO STRING(255);
END_VAR
END_METHOD

METHOD PRVWRITEUSER : BOOL
VAR_INPUT
	PVUMUSER : POINTER TO VUM_User;
	DWFILE : SysFile.RTS_IEC_HANDLE;
	BEMPTYPASSWORDALLOWED : BOOL;
END_VAR
END_METHOD

METHOD PRVWRITEVALUE : BOOL
VAR_INPUT
	PDATA : POINTER TO BYTE;
	DWSIZE : DWORD;
	DWFILE : SysFile.RTS_IEC_HANDLE;
END_VAR
END_METHOD

(* ---- VISUUSERMGMTCYCLICCALL.fb ---- *)
FUNCTION_BLOCK VISUUSERMGMTCYCLICCALL
VAR
	_BINIT : BOOL := TRUE;
	_NCOUNTER : INT;
	_CLIENTLISTENER : VisuFbClientManagerListener;
	M_ITFCLIENTMANAGERLISTENER : VisuElems.IClientManagerListener := _ClientListener;
	_DIALOGLISTENER : VisuUserMgmtDialogManagerListener;
	M_ITFDIALOGMANAGERLISTENER : VisuElems.IDialogManagerListener := _DialogListener;
END_VAR
END_FUNCTION_BLOCK

METHOD CYCLICCALL : BOOL
END_METHOD

(* ---- VISUUSERMGMTDIALOGMANAGERLISTENER.fb ---- *)
FUNCTION_BLOCK VISUUSERMGMTDIALOGMANAGERLISTENER
END_FUNCTION_BLOCK

METHOD CLOSEDIALOG
VAR_INPUT
	PCLIENTDATA : POINTER TO VisuElems.VisuStructClientData;
	ITFDIALOG : VisuElems.IVisualisationDialog;
	BALLCLIENTDIALOGSCLOSED : BOOL;
	BMODAL : BOOL;
END_VAR
END_METHOD

METHOD OPENDIALOG
VAR_INPUT
	PCLIENTDATA : POINTER TO VisuElems.VisuStructClientData;
	ITFDIALOG : VisuElems.IVisualisationDialog;
	BMODAL : BOOL;
END_VAR
END_METHOD

(* ---- VISUUSERMGMTFBLOGINLOCKOUTTIMEINFOVECTOR.fb ---- *)
FUNCTION_BLOCK VISUUSERMGMTFBLOGINLOCKOUTTIMEINFOVECTOR EXTENDS VisuFbBaseVector
VAR
	_PENTRIES : POINTER TO VUM_StructLoginLockoutTimeUserEntry;
END_VAR
END_FUNCTION_BLOCK

METHOD ADDENTRY : UDINT
VAR_INPUT
	WSTUSERNAME : WSTRING;
	DWLOCKOUTSTART : DWORD;
	BUSEADMINLOCKOUTTIME : BOOL;
END_VAR
END_METHOD

METHOD GETINDEXOFUSERENTRY : DINT
VAR_INPUT
	WSTUSER : WSTRING;
END_VAR
END_METHOD

METHOD GETUSERENTRY : POINTER TO VUM_StructLoginMaxAttemptsUserEntry
VAR_INPUT
	WSTUSER : WSTRING;
END_VAR
END_METHOD

METHOD ABSTRASSIGN : UDINT
VAR_INPUT
	PBT : POINTER TO BYTE;
	UDIINDEX : UDINT;
END_VAR
END_METHOD

METHOD ABSTRDATAPTRCHANGED : UDINT
END_METHOD

METHOD ABSTRGETELEMENTPTR : UDINT
VAR_INPUT
	UDIINDEX : UDINT;
END_VAR
VAR_OUTPUT
	PENTRY : POINTER TO BYTE;
END_VAR
END_METHOD

METHOD ABSTRSIZEOFELEMENT : UDINT
END_METHOD

(* ---- VISUUSERMGMTFBLOGINMAXATTEMPTSINFOVECTOR.fb ---- *)
FUNCTION_BLOCK VISUUSERMGMTFBLOGINMAXATTEMPTSINFOVECTOR EXTENDS VisuFbBaseVector
VAR
	_PENTRIES : POINTER TO VUM_StructLoginMaxAttemptsUserEntry;
END_VAR
END_FUNCTION_BLOCK

METHOD ADDENTRY : UDINT
VAR_INPUT
	WSTUSERNAME : WSTRING;
	USILOGINATTEMPTS : USINT;
END_VAR
END_METHOD

METHOD GETINDEXOFUSERENTRY : DINT
VAR_INPUT
	WSTUSER : WSTRING;
END_VAR
END_METHOD

METHOD GETUSERENTRY : POINTER TO VUM_StructLoginMaxAttemptsUserEntry
VAR_INPUT
	WSTUSER : WSTRING;
END_VAR
END_METHOD

METHOD ABSTRASSIGN : UDINT
VAR_INPUT
	PBT : POINTER TO BYTE;
	UDIINDEX : UDINT;
END_VAR
END_METHOD

METHOD ABSTRDATAPTRCHANGED : UDINT
END_METHOD

METHOD ABSTRGETELEMENTPTR : UDINT
VAR_INPUT
	UDIINDEX : UDINT;
END_VAR
VAR_OUTPUT
	PENTRY : POINTER TO BYTE;
END_VAR
END_METHOD

METHOD ABSTRSIZEOFELEMENT : UDINT
END_METHOD

(* ---- VISUUSERMGMTPROVIDER.fb ---- *)
FUNCTION_BLOCK VISUUSERMGMTPROVIDER
VAR
	ARRUSERSTODISPLAY : ARRAY [0..(MAX_VISIBLE_USERS - 1)] OF VUM_UserInternal;
	ARRUSERSTODISPLAYMAIN : POINTER TO VUM_UserInternal;
	ARRUSERSTODISPLAYMAINSZ : UDINT := MAX_VISIBLE_USERS;
	VMUSER : VUM_User;
	ARRGROUPSELECTION : ARRAY [0..MAX_USER_GROUPS] OF VUM_GroupSelection;
	IMAXGROUPS : INT := -1;
	LASTSELECTEDUSER : VUM_UserInternal;
	LASTEDITEDUSER : VUM_UserInternal;
	UDIUSERCOUNT2 : UDINT;
	UDIGROUPPOS : UDINT;
	UDIPOS : UDINT;
	UDILASTPOS : UDINT;
	UDISELECTION : UDINT := INVALID_SELECTION_OR_POS;
	UDILASTSELECTION : UDINT := INVALID_SELECTION_OR_POS;
	DWDIALOGRESULTOK : BOOL;
	DWLASTDIALOGRESULTOK : BOOL;
	DWDIALOGRESULTCANCEL : BOOL;
	DWLASTDIALOGRESULTCANCEL : BOOL;
	STUSERNAME : WSTRING;
	STFULLNAME : WSTRING;
	STPASSWORD : WSTRING;
	STACKNOWLEDGEPASSWORD : WSTRING;
	BDEACTIVATED : BOOL;
	BCHGPASSFIRSTLOGIN : BOOL;
	BINSERTUSER : BOOL;
	BREMOVEUSER : BOOL;
	BRESULT : BOOL;
	DWRESULT : DWORD;
	UDILASTERROR : UDINT;
	BPREVENTDELETINGLASTADMIN : BOOL;
	BRTSBASED : BOOL;
	BHEADERINVIS : BOOL;
	BDELETEINVIS : BOOL;
	IMOVEX : INT;
	IMOVEY : INT;
	BGRPSKO : BOOL;
	ITFVISUUSERMGMT : IVisuUserMgmt;
	ITFVISUUSERMGMT4 : IVisuUserMgmt4;
	_UDIUSERCOUNT : UDINT;
	_UDIRESULTVERSION : UDINT;
	_XSWAPPINGNEEDED : BOOL;
	_VISUUSERMGMTSTATE : EVisuUserMgmtState;
	_PCLIENTDATA : POINTER TO VisuElems.VisuStructClientData;
	_BCURRENTSTATE : BYTE := 0;
	_BLASTCURRENTSTATE : BYTE := 0;
	_DWUSERDB : DWORD;
	_BCANCLOSE : BOOL;
	_IINDEXARRAY : INT;
	_IINDEX : INT;
	_WSTADMINNAME : WSTRING(79);
	_EEDITTYPE : VUM_EditType;
	VUMP_STATE_NONE : BYTE := 0;
	VUMP_STATE_GET_USER_DB : BYTE := 1;
	VUMP_STATE_EDIT_USER : BYTE := 2;
	VUMP_STATE_RELOAD_USER_LIST : BYTE := 3;
	VUMP_STATE_GET_USER_COUNT : BYTE := 4;
	VUMP_STATE_GET_USERS : BYTE := 5;
	VUMP_STATE_SEND_USER_BEFOR_CLOSE : BYTE := 6;
	VUMP_STATE_SET_USER_DB : BYTE := 7;
	VUMP_STATE_TIMEOUT : DWORD := 2000;
END_VAR
END_FUNCTION_BLOCK

METHOD INITIALIZE : BOOL
VAR_INPUT
	IVISUUSERMGMT : IVisuUserMgmt;
	PCLIENTDATA : POINTER TO VisuElems.VisuStructClientData;
END_VAR
END_METHOD

METHOD SETEXTUSERSTODISPLAYARRAY : INT
VAR_INPUT
	ARR : POINTER TO VUM_UserInternal;
	ARRSIZE : UDINT;
END_VAR
END_METHOD

METHOD SETUSERCOUNT : BOOL
VAR_INPUT
	UDIUSERCOUNT : UDINT;
END_VAR
END_METHOD

METHOD SETUSERDB : BOOL
VAR_INPUT
	UDIUSERDB : UDINT;
END_VAR
END_METHOD

METHOD SETUSERS : BOOL
VAR_INPUT
	UDIUSERCOUNT : UDINT;
	PARRUSERS : POINTER TO ARRAY [0..(MAX_VISIBLE_USERS - 1)] OF VUM_User;
END_VAR
END_METHOD

METHOD PRVCHANGEUSERLEGACY : BOOL
VAR_INPUT
	DWUSERDB : DWORD;
	PVUMUSER : POINTER TO VUM_UserInternal;
	UDIINDEX : UDINT;
	EEDITTYPE : VUM_EditType;
END_VAR
END_METHOD

METHOD PRVCHECKANDSENDUSER : BOOL
VAR_OUTPUT
	BCANCLOSE : BOOL;
END_VAR
END_METHOD

METHOD PRVCHECKUSERISADMIN : BOOL
VAR_INPUT
	PVUMUSER : POINTER TO VUM_UserInternal;
	ITFVISUUSERMGMT : IVisuUserMgmt;
END_VAR
END_METHOD

METHOD PRVCMPUSER : BOOL
VAR_INPUT
	PVUMUSER1 : POINTER TO VUM_UserInternal;
	PVUMUSER2 : POINTER TO VUM_UserInternal;
END_VAR
END_METHOD

METHOD PRVFILLUSER : BOOL
VAR_INPUT
	PVUMUSERIN : POINTER TO VUM_UserInternal;
	BTOTEXTFIELDS : BOOL;
END_VAR
END_METHOD

METHOD PRVGETUSERSLEGACY : DWORD
VAR_INPUT
	DWUSERDB : DWORD;
	UDISTARTINDEX : UDINT;
	UDIENDINDEX : UDINT;
	PARR : POINTER TO ARRAY [0..10] OF VUM_UserInternal;
	UDIARRSIZE : UDINT;
END_VAR
END_METHOD

METHOD PRVISCURRENTUSERADMIN : BOOL
VAR_INPUT
	PVUMUSER : POINTER TO VUM_UserInternal;
END_VAR
END_METHOD

METHOD PRVSENDUSER : BOOL
VAR_INPUT
	EEDITTYPE : VUM_EditType;
	BCHECKFOREMPTYPASSWORD : BOOL;
END_VAR
END_METHOD

METHOD PRVSETCURRENTADMINUSER : BOOL
VAR_INPUT
	PVUMUSER : POINTER TO VUM_UserInternal;
END_VAR
END_METHOD

METHOD PRVSETNEWUSERDB : BOOL
VAR_INPUT
	DWUSERDB : DWORD;
	BRESULTOK : BOOL;
END_VAR
END_METHOD

(* ---- VISUUSERMGMTSEM.fb ---- *)
FUNCTION_BLOCK VISUUSERMGMTSEM
VAR
	_HSEM : SysTypes.RTS_IEC_HANDLE;
END_VAR
END_FUNCTION_BLOCK

METHOD ENTER
END_METHOD

METHOD FB_EXIT : BOOL
VAR_INPUT
	BINCOPYCODE : BOOL;
END_VAR
END_METHOD

METHOD FB_INIT
VAR_INPUT
	BINITRETAINS : BOOL;
	BINCOPYCODE : BOOL;
END_VAR
END_METHOD

METHOD LEAVE
END_METHOD
